FUNCTION_BLOCK MoveRelativeTask EXTENDS TcoCore.TcoTask IMPLEMENTS ITcoDriveSimple
VAR
    {attribute addProperty Name "<#Distance#>"}
    _distance : LREAL;
    {attribute addProperty Name "<#Velocity#>"}
    _velocity : LREAL;
    {attribute addProperty Name "<#Acceleration#>"}
    _acceleration : LREAL;
    {attribute addProperty Name "<#Deceleration#>"}
    _deceleration : LREAL;
    {attribute addProperty Name "<#Jerk#>"}
    _jerk : LREAL;
END_VAR
VAR
    {attribute 'hide'}
    _axisRef : REFERENCE TO TcoAxisRef;
    {attribute 'hide'}
    _mcMoveRelative : Tc2_MC2.MC_MoveRelative;
    {attribute 'hide'}
    _dummyPreconditionOK : BOOL;
END_VAR

IF NOT __ISVALIDREF(_axisRef) THEN
    IF __ISVALIDREF(DriveRef) THEN
        _axisRef REF= DriveRef.AxisRef;
    ELSE
        RETURN;
    END_IF
END_IF
IF Execute() THEN
    _dummyPreconditionOK := TRUE;

    IF NOT DriveRef._movementState.MovePreconditionsOk(THIS^, _dummyPreconditionOK) THEN
        Messenger.Error('To be implemented');
        RETURN;
    END_IF

    _mcMoveRelative(Axis := _axisRef,
        Execute := NOT _mcMoveRelative.Busy,
        Distance := _distance,
        Velocity := _velocity,
        Acceleration := _acceleration,
        Deceleration := _deceleration,
        Jerk := _jerk,
        BufferMode := Tc2_MC2.MC_Aborting,
        Done =>,
        Busy =>,
        Active =>,
        CommandAborted =>,
        Error =>,
        ErrorID =>);

    IF _mcMoveRelative.CommandAborted THEN
        THIS^.Abort();
    END_IF

    DoneWhen(_mcMoveRelative.Done);
    ThrowWhen(_mcMoveRelative.Error);

END_IF

PROPERTY DriveRef : REFERENCE TO TcoDriveSimple
GET
VAR
    _drive : ITcoDriveSimple := 0;
END_VAR
IF __QUERYINTERFACE(THIS^.Parent, _drive) THEN
    DriveRef REF= _drive.DriveRef;
END_IF
END_GET
END_PROPERTY

METHOD PUBLIC FB_init : BOOL
VAR_INPUT
    bInitRetains : BOOL; // if TRUE, the retain variables are initialized (warm start / cold start)
    bInCopyCode : BOOL; // if TRUE, the instance afterwards gets moved into the copy code (online change)
  	ParentObject : ITcoObject;	
END_VAR
END_METHOD

METHOD INTERNAL InvokeWithParams : ITcoTaskStatus
VAR_INPUT
    inDistance : LREAL;
    inVelocity : LREAL;
    inAcceleration : LREAL;
    inDeceleration : LREAL;
    inJerk : LREAL;
END_VAR
_distance := inDistance;
_velocity := inVelocity;
_acceleration := inAcceleration;
_deceleration := inDeceleration;
_jerk := inJerk;
InvokeWithParams := THIS^.Invoke();
END_METHOD

(*~
	<docu>
		<summary>
			Executes when task is aborted.
		</summary>			
	</docu>	
~*)
METHOD PROTECTED OnAbort
IF NOT __ISVALIDREF(_axisRef) THEN
    IF __ISVALIDREF(DriveRef) THEN
        _axisRef REF= DriveRef.AxisRef;
    ELSE
        RETURN;
    END_IF
END_IF

THIS^.DriveRef.Stop(-1, -1);
THIS^.DriveRef._movementState.Restore();
_mcMoveRelative(Axis := _axisRef, Execute := FALSE);
END_METHOD

(*~
	<docu>
		<summary>
			Executes when task reaches the ```Done``` state .
		</summary>			
	</docu>	
~*)
METHOD PROTECTED OnDone
THIS^.DriveRef._movementState.Restore();
_mcMoveRelative(Axis := _axisRef, Execute := FALSE);
END_METHOD

(*~
	<docu>
		<summary>
			Executes when task reaches the ```Error``` state.
			<para>
				Do not confuse with <see cref="PlcDocu.TcoCore.TcoTask.WhileError()"/>, that is called cyclically until '''Error''' state is left.
			</para>
		</summary>			
	</docu>	
~*)
METHOD PROTECTED OnError
THIS^.DriveRef._movementState.Restore();
IF NOT _axisRef.Status.Error THEN
	DriveRef.SetErrorID(DriveRef._moveRelativeTask._mcMoveRelative.ErrorID);
END_IF
_mcMoveRelative(Axis := _axisRef, Execute := FALSE);
END_METHOD

METHOD PROTECTED OnStart
_mcMoveRelative(Axis := _axisRef, Execute := FALSE);
END_METHOD

(*~
	<docu>
		<summary>
			Restores this instance to the Ready state. Can be called explicitly or from within one of the restore mechanisms.
			<para>
				See also <see cref="PlcDocu.TcoCore.TcoTask.AutoRestorable()"/>
			</para>
		</summary>			
	</docu>	
~*)
METHOD Restore : ITcoRestorable
SUPER^.Restore();
END_METHOD

(*~
	<docu>
		<summary>
			Executes until task is in ```Error``` state .
		</summary>			
	</docu>	
~*)
METHOD PROTECTED WhileError
IF NOT _axisRef.Status.Error THEN
	DriveRef.SetErrorID(DriveRef._moveRelativeTask._mcMoveRelative.ErrorID);
    _mcMoveRelative(Axis := _axisRef, Execute := FALSE);
END_IF
END_METHOD

END_FUNCTION_BLOCK

(* stored: Version 1.1.0.1, ProductVersion 3.1.4024.12
   POU MoveRelativeTask: Id {ab769f25-b35b-017a-34f4-12fb5831bde5}, SpecialFunc None
   Property DriveRef: Id {146efb26-7f32-04da-32b9-93685dec6a03}
   Get Get: Id {190a9f73-0399-046c-1c21-3bcf8e4250e7}
   Method FB_init: Id {aa0a4a5c-48ac-02d1-3cc2-173990343fe1}
   Method InvokeWithParams: Id {01411d53-ac5f-0768-12a4-5b448e2f644f}
   Method OnAbort: Id {b2c16ee0-afd5-068f-3960-07dec1b46405}
   Method OnDone: Id {57a9f802-273a-0f02-25dc-2e184a738dba}
   Method OnError: Id {04568080-7829-0dc8-1387-20a80a858f6e}
   Method OnStart: Id {3ab86d75-bbf1-0431-304b-74df4f8dfd95}
   Method Restore: Id {e976de80-cfea-01a1-1fd9-673984f12c06}
   Method WhileError: Id {5b8e54de-475c-0f46-2d99-ccc66c7867aa} *)
